FUNCTION_BLOCK FB_MunschExtruderAir_1
(*

The function block used to control air pressure.

Constructor: 		Patryk Panylo
Company:		E. Riexinger GmbH
Date:			04.11.2016
Version:			1.00

Date:			Revision:		Who:				Comment
dd.mm.yyyy		x.xx			Initials			comment

*)
VAR_INPUT
	(* Input variables / Eingang Variablen *)
	bEnable					:BOOL;						(* Enable FB signal *)
	bIn						:BOOL;						(* Input signal *)
	bExtruderAirOn			:BOOL;						(* Extruder air on *)
	tAirOk					:TIME := t#5s;					(* Timer to delay output air ok *)
	tAirOff					:TIME := t#5s;					(* Timer to delay output air off *)
	tTimeOut					:TIME := t#5s;					(* Timeout *)
END_VAR
VAR_OUTPUT
	(* Output variables / Ausgang Variablen *)
	bAirOk					:BOOL;						(* Air pressure ok *)
	bAirOn					:BOOL;						(* Air pressure on *)
	bError					:BOOL;						(* Error by no air pressure *)
	udnErrorNo				:UDINT;
	udnMessageNo			:UDINT;
END_VAR
VAR
	(* Enummerations *)

	(* Variables *)

	(* References *)

	(* Interfaces *)

	(* Instances *)
	tonDelayAirOk				:TON;						(* Timer to delay *)
	tofDelayAirOff					:TOF;						(* Timer to delay *)
	fbExtrudingAir					:FB_AirPressure;
END_VAR


IF NOT bEnable
THEN
	fbExtrudingAir(
		bEnable := FALSE
	);

	bAirOk := FALSE;
	RETURN;
END_IF

fbExtrudingAir(
	bEnable := bEnable,
	bIn := bIn,
	bNoEStop := bExtruderAirOn,
	tTimeOut := tTimeOut,
	bError => bError,
	udnErrorNo => udnErrorNo,
	udnMessageNo => udnMessageNo
);

tonDelayAirOk(
	IN := fbExtrudingAir.bOut,
	PT := tAirOk
);

bAirOk := tonDelayAirOk.Q;

tofDelayAirOff(
	IN := fbExtrudingAir.bAirOn,
	PT := tAirOff
);

bAirOn := tofDelayAirOff.Q;

END_FUNCTION_BLOCK

(* stored: Version 1.1.0.1, ProductVersion 3.1.4024.15
   POU FB_MunschExtruderAir_1: Id {9a34f482-e02e-4813-b61b-d2ec53884544}, SpecialFunc None *)
